(* IEC 61131-3 sources: trust-platform/editors/vscode/src/test/fixtures/control-studio-engineer/src, 1 file *)

(* ---- Main.st ---- *)
PROGRAM Main
VAR
    Kp : LREAL := LREAL#1.0;
    Manual : BOOL := TRUE;
    ManualCommand AT %ML8 : LREAL := LREAL#0.0;
    SP AT %ML0 : LREAL := LREAL#0.0;
    PV AT %IL0 : LREAL;
    MV AT %QL0 : LREAL;
END_VAR

IF Manual THEN
    MV := ManualCommand;
ELSE
    MV := LIMIT(LREAL#-20.0, Kp * (SP - PV), LREAL#20.0);
END_IF;
END_PROGRAM

CONFIGURATION Config
RESOURCE Res ON PLC
    TASK MainTask(INTERVAL := T#20ms, PRIORITY := 1);
    PROGRAM Main WITH MainTask : Main;
END_RESOURCE
END_CONFIGURATION
